// TwinCAT 3 PLC project DaisyChain
// ProgramVersion: 3.1.4023.0
// libraries:
//   Tc2_Standard, * (Beckhoff Automation GmbH)
//   Tc2_System, * (Beckhoff Automation GmbH)
//   Tc3_Module, * (Beckhoff Automation GmbH)
// project tree:
//   DUTs/ EthercatDevice.TcDUT
//   / PlcTask.TcTTO
//   POUs/ MAIN.TcPOU
// real-time tasks:
//   TASK PlcTask: cycle T#10ms, priority 20, ADS port 350

CONFIGURATION DaisyChain
    RESOURCE PLC ON TwinCAT3
        TASK PlcTask(INTERVAL := T#10ms, PRIORITY := 20);
        PROGRAM MAIN WITH PlcTask : MAIN;
    END_RESOURCE
END_CONFIGURATION

// ---- DUTs/EthercatDevice.TcDUT
TYPE EthercatDevice :
STRUCT
	dir : BYTE ;
	speed : WORD ;
	dummyDataOut AT %Q*: DWORD ;
	dummyDataIn AT %I*: DWORD ;
END_STRUCT
END_TYPE

// ---- POUs/MAIN.TcPOU
PROGRAM MAIN

VAR CONSTANT 
    deviceCount : WORD := 3;
END_VAR

VAR
	{attribute 'TcLinkTo' := '[1].dummyDataOut := TIID^Device_1^Box 1 (sample_app)^Outputs process data mapping^Trigger;
							[1].dummyDataIn := TIID^Device_1^Box 1 (sample_app)^Inputs process data mapping^Counter;
							[2].dummyDataOut := TIID^Device_1^Box 2 (sample_app)^Outputs process data mapping^Trigger;
							[2].dummyDataIn := TIID^Device_1^Box 2 (sample_app)^Inputs process data mapping^Counter;
							[3].dummyDataOut := TIID^Device_1^Box 3 (sample_app)^Outputs process data mapping^Trigger;
							[3].dummyDataIn := TIID^Device_1^Box 3 (sample_app)^Inputs process data mapping^Counter'}
	device : ARRAY [1..deviceCount] OF EthercatDevice ;
	counter: WORD;
END_VAR

FOR counter:=1 TO deviceCount BY 1 DO

    device[counter].dummyDataOut:= SHL(device[counter].dir,2*8) OR device[counter].speed ;

END_FOR;

END_PROGRAM
